// TIA Portal V21 export
// export: Created 2026-11-07T00:00:00Z, ExportSetting WithDefaults
TextList "TL_State"  ListRange=Range
  TextListEntry   Text="OFF"
  TextListEntry   From=1, To=1, Text="INIT"
